(* Processor test double that retains one emitted record for assertions. *)
FUNCTION_BLOCK FB_LogRecordProcessor_ForRecordInspection EXTENDS FB_LogRecordProcessor_Simple
VAR_OUTPUT
	record: POINTER TO FB_LogRecord;
	lastOperationSucceeded: BOOL := FALSE;
	failureResult: E_LogRecordCloneFailureReason;
END_VAR

METHOD free
IF THIS^.record <> 0 THEN
	THIS^.record^.delete(pSelf:=THIS^.record);
END_IF
END_METHOD

METHOD onEmit
VAR_INPUT
	logRecord: REFERENCE TO FB_LogRecord;
END_VAR
THIS^.free();
THIS^.lastOperationSucceeded := logRecord.cloneTo(
	pDest:=THIS^.record,
	failureReason=>THIS^.failureResult
);
END_METHOD

METHOD pop : POINTER TO FB_LogRecord
pop := THIS^.record;
THIS^.record := 0;
END_METHOD

END_FUNCTION_BLOCK

(* stored: Version 1.1.0.1
   POU FB_LogRecordProcessor_ForRecordInspection: Id {86e0c01f-365f-4c34-a5f8-f56ecceaf360}, SpecialFunc None
   Method free: Id {9d6f0dd6-04e2-43c1-b207-46bd50021591}
   Method onEmit: Id {60b935aa-5fef-4d49-a6b2-6e0283d21352}
   Method pop: Id {3930a8d2-bfba-4caf-bbd7-c6b54b336880} *)
